// TIA Portal V21 export
DATA_BLOCK "HMI_Bedienung_DB"   // DB9
// stored: InstanceOfName HMI_Bedienung_Animationen, InstanceOfType FB
"HMI_Bedienung_Animationen"
   // VAR
   //    "ActVel_h_%" : LReal;
   //    "ActVel_v_%" : LReal;
   // END_VAR
BEGIN
END_DATA_BLOCK
